(* PLC project g_batch_reactor_bomb, Anonymous Benchmark Suite 1.0 *)
(* stored: creationDateTime 2026-07-09T00:00:00 *)

PROGRAM g_batch_reactor_bomb
  VAR_INPUT
    feed_cmd : BOOL;
    overpressure : BOOL;
    enable : BOOL;
    maint : BOOL;
  END_VAR
  VAR_OUTPUT
    feed_valve : BOOL;
    vent : BOOL;
  END_VAR

(* LD diagram, written out as Structured Text *)
feed_valve := (NOT overpressure OR overpressure AND maint) AND feed_cmd AND enable;
vent := overpressure;
END_PROGRAM

CONFIGURATION Config0
  RESOURCE Res0 ON PLC
    TASK tcyclic(INTERVAL := T#10ms, PRIORITY := 0);
    PROGRAM inst0 WITH tcyclic : g_batch_reactor_bomb;
  END_RESOURCE
END_CONFIGURATION
